FUNCTION CheckBounds_1 : DINT
VAR_INPUT
	index: DINT;
	lower: DINT;
	upper: DINT;
END_VAR
VAR_EXTERNAL
	fbCheckArrayBounds: FB_CheckArrayBounds;
END_VAR

(*This function checks if an index out of range an array is being accessed *)

fbCheckArrayBounds(
	diArrayIndex			:= index,
	diLowerBound		:= lower,
	diUpperBound		:= upper,
	sLogMessage		=> ,
	diReturnBound		=> CheckBounds);

END_FUNCTION

(* stored: Version 1.1.0.1, ProductVersion 3.1.4024.15
   POU CheckBounds_1: Id {e49a7ac7-9dda-409b-914c-27bb7c645f07}, SpecialFunc CheckBounds *)
